// TIA Portal V19 export
// export: Created 2026-01-15T10:00:00.0000000Z, ExportSetting WithReadOnly
ORGANIZATION_BLOCK "Main"   // OB1, LAD, Example_ProgramCycle
// stored: AutoNumber false, IsKnowHowProtected false, ModifiedDate 2026-01-10T09:00:00.0000000Z, PriorityNumber 1
   VAR_INPUT
      Initial_Call : Bool;
   END_VAR
BEGIN

REGION Network 1: Run permissive
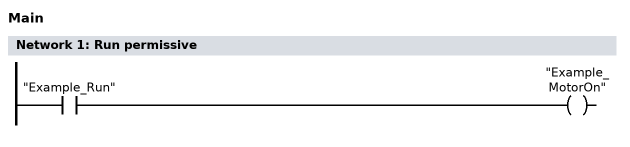
   RUNG wire#powerrail
      Contact( "Example_Run" )
      Coil( "Example_MotorOn" )
   END_RUNG
   // the same network as SCL:
   "Example_MotorOn" := "Example_Run";
END_REGION

REGION Network 2 (SCL): Speed handling
   "DB_ExampleData".Speed := "Example_Speed";
   "FC_ExampleScale"(In := "Example_Speed", Out => "DB_ExampleData".Scaled);
END_REGION
END_ORGANIZATION_BLOCK
